Staubli VAL3: appStart.dtx

public string sAppName = "MainApp"
public string sDbId = ""
public string sRobotModel
public string sRobotSN
public string sCtrlSN
public string sProfile
public string sProfileRaw
public string sLogin[2]
  [0] = "operator"
  [1] = "programmer"
public string sRoleName[2]
  [0] = "生产员"
  [1] = "工程师"
public bool bFunc[9]
public string sFuncBg[9]
  [0] = "#DCDCDC"
  [1] = "#DCDCDC"
  [2] = "#DCDCDC"
  [3] = "#DCDCDC"
  [4] = "#DCDCDC"
  [5] = "#DCDCDC"
  [6] = "#DCDCDC"
  [7] = "#DCDCDC"
  [8] = "#DCDCDC"
public bool bBtnPressed[9]
